(* IEC 61131-3 sources: ST2CPP/examples/projects/syntax_tests, 37 files *)

(* ---- __combined.st ---- *)
(* test_class.st — CLASS 和方法调用测试 *)

CLASS MATH_HELPER
    VAR
        LAST_RESULT : DINT;
        CALL_COUNT  : INT;
    END_VAR

    METHOD ADD : DINT
        VAR_INPUT
            A : DINT;
            B : DINT;
        END_VAR
        LAST_RESULT := A + B;
        CALL_COUNT := CALL_COUNT + 1;
        ADD := LAST_RESULT;
    END_METHOD

    METHOD SUBTRACT : DINT
        VAR_INPUT
            A : DINT;
            B : DINT;
        END_VAR
        LAST_RESULT := A - B;
        CALL_COUNT := CALL_COUNT + 1;
        SUBTRACT := LAST_RESULT;
    END_METHOD

    METHOD GET_COUNT : INT
        GET_COUNT := CALL_COUNT;
    END_METHOD
END_CLASS

PROGRAM TEST_CLASS
    VAR
        Helper      : MATH_HELPER;
        R1          : DINT;
        R2          : DINT;
        Count       : INT;
    END_VAR

    R1 := Helper.ADD(10, 20);
    ASSERT(R1 = 30);

    R2 := Helper.SUBTRACT(50, 15);
    ASSERT(R2 = 35);

    Count := Helper.GET_COUNT();
    ASSERT(Count = 2);

    ASSERT(TRUE);
END_PROGRAM

(* test_class_minimal.st — 最小 CLASS 测试 *)

CLASS BASE_CTRL
    VAR
        BASE_STATE : INT := 0;
    END_VAR

    METHOD GET_VALUE : INT
        GET_VALUE := BASE_STATE;
    END_METHOD
END_CLASS

PROGRAM TEST_MINIMAL
    VAR
        Ctrl : BASE_CTRL;
        R    : INT := 0;
    END_VAR
    R := Ctrl.GET_VALUE();
END_PROGRAM

(* test_class_no_extend.st — CLASS 无继承测试 *)

CLASS MY_CLASS
    VAR
        DATA : INT := 0;
    END_VAR

    METHOD GET_DATA : INT
        GET_DATA := DATA;
    END_METHOD
END_CLASS

PROGRAM TEST_NO_EXTEND
    VAR
        Obj : MY_CLASS;
        R   : INT := 0;
    END_VAR
    R := Obj.GET_DATA();
END_PROGRAM

TYPE MyStruct :
STRUCT
    X : INT;
    Y : INT;
END_STRUCT;
END_TYPE

PROGRAM AT_STRUCT
  VAR_INPUT
    Raw AT %ID0 : MyStruct;
  END_VAR
  VAR_OUTPUT
    Out AT %QD0 : MyStruct;
  END_VAR
  VAR
    LocalX : INT;
  END_VAR
    LocalX := Raw.X;
    Out.Y := Raw.X + 1;
END_PROGRAM

FUNCTION_BLOCK TEST_FB
    VAR_INPUT
        X : INT;
    END_VAR
    VAR_OUTPUT
        Y : INT;
    END_VAR
    VAR
        S : INT := 0;
    END_VAR

    CASE S OF
        0:
            Y := 16#0007;
            IF X > 0 THEN
                S := 1;
            END_IF;
        1:
            Y := 16#000F;
            S := 0;
        ELSE
            Y := 0;
    END_CASE;
END_FUNCTION_BLOCK

PROGRAM IO_TEST
  VAR_INPUT
    BitInput AT %IX1.3 : BOOL;
    ByteInput AT %IB5 : USINT;
    WordInput AT %IW2 : INT;
    DWordInput AT %ID1 : DINT;
  END_VAR
  VAR_OUTPUT
    BitOutput AT %QX0.7 : BOOL;
    ByteOutput AT %QB10 : USINT;
    WordOutput AT %QW3 : INT;
    DWordOutput AT %QD2 : DINT;
  END_VAR
  VAR
    Temp : INT;
    Result : INT;
  END_VAR
    Temp := WordInput + 5;
    IF BitInput THEN
        BitOutput := TRUE;
    ELSE
        BitOutput := FALSE;
    END_IF;
    ByteOutput := ByteInput;
    WordOutput := Temp;
    DWordOutput := DWordInput * 2;
    Result := WordInput * 10;
END_PROGRAM

PROGRAM IO_READBACK
  VAR_INPUT
    Cmd AT %IX0.0 : BOOL;
  END_VAR
  VAR_OUTPUT
    OutVal AT %QW2 : INT;
    OutFlag AT %QX0.1 : BOOL;
  END_VAR
  VAR
    Readback : INT;
    FlagCopy : BOOL;
  END_VAR
    OutVal := 42;
    OutFlag := Cmd;
    Readback := OutVal;
    FlagCopy := OutFlag;
END_PROGRAM

PROGRAM AT_VAR
  VAR
    MyInput AT %IW2 : INT;
    MyOutput AT %QW1 : INT;
    MyFlag AT %QX0.5 : BOOL;
  END_VAR
    MyOutput := MyInput * 2;
    IF MyInput > 100 THEN
        MyFlag := TRUE;
    ELSE
        MyFlag := FALSE;
    END_IF;
END_PROGRAM

(* test_bitwise.st — 测试 Bug 3: AND/OR 对非 BOOL 操作数
 *
 * 问题：VisitAnd_expr 强制要求 BOOL 类型，拒绝 INT 操作数
 * 预期：AND/OR 应支持 ANY_BIT 多态（BYTE/WORD/DWORD/INT 等）
 *       编译器 mapOperator 已将 AND→&, OR→|，只需放宽静态检查
 *)

PROGRAM TEST_BITWISE
    VAR
        A     : INT := 16#FF00;
        B     : INT := 16#0F0F;
        MASK  : INT := 16#00FF;
        AND_R : INT := 0;
        OR_R  : INT := 0;
        XOR_R : INT := 0;
    END_VAR

    AND_R := A AND MASK;
    OR_R  := A OR B;
    XOR_R := A XOR B;

    ASSERT(AND_R = 16#0000);
    ASSERT(OR_R = 16#FF0F);
    ASSERT(XOR_R = 16#F0F0);
END_PROGRAM

FUNCTION_BLOCK MY_FB
    VAR_INPUT X : INT; END_VAR
    VAR_OUTPUT Y : INT; END_VAR
    Y := X + 1;
END_FUNCTION_BLOCK

PROGRAM TEST_FB_ARR
    VAR
        Fbs : ARRAY[0..2] OF MY_FB;
        I : INT;
    END_VAR
    FOR I := 0 TO 2 DO
        Fbs[I](X := I);
    END_FOR;
END_PROGRAM

(* test_fb_output.st — 测试 FB 输出参数 => 在 update 后读回
 *
 * 问题：FB 调用时 => 参数在 update() 后没有从 FB 实例读回
 * 预期：SM(STATUS => MyStatus) 应在 update 后将 FB 的 STATUS 字段读回 MyStatus
 *)

FUNCTION_BLOCK STATE_MACHINE
    VAR_INPUT
        CMD : INT;
    END_VAR
    VAR_OUTPUT
        STATUS : INT;
        DONE   : BOOL;
    END_VAR
    VAR
        MODE : INT := 0;
    END_VAR

    CASE CMD OF
        0:
            MODE := 0;
            STATUS := 0;
            DONE := FALSE;
        1:
            MODE := 1;
            STATUS := 10;
            DONE := TRUE;
        2:
            MODE := 2;
            STATUS := 20;
            DONE := TRUE;
    END_CASE
END_FUNCTION_BLOCK

PROGRAM TEST_FB_OUTPUT
    VAR
        SM       : STATE_MACHINE;
        MyStatus : INT := 0;
        MyDone   : BOOL := FALSE;
    END_VAR

    SM(CMD := 1, STATUS => MyStatus, DONE => MyDone);
    ASSERT(MyStatus = 10);
    ASSERT(MyDone = TRUE);

    SM(CMD := 2, STATUS => MyStatus, DONE => MyDone);
    ASSERT(MyStatus = 20);
    ASSERT(MyDone = TRUE);

    SM(CMD := 0, STATUS => MyStatus, DONE => MyDone);
    ASSERT(MyStatus = 0);
    ASSERT(MyDone = FALSE);
END_PROGRAM

(* test_fc_return.st — 测试 Bug 1: FC 末尾多余 return;
 *
 * 问题：TranslateReturn 对非 void FC 也输出 return; 导致编译报错
 * 预期：非 void FC 应该 return <returnValue>; 而不是 return;
 *)

FUNCTION ADD : DINT
    VAR_INPUT
        A : DINT;
        B : DINT;
    END_VAR
    ADD := A + B;
END_FUNCTION

FUNCTION CLAMP : DINT
    VAR_INPUT
        VAL  : DINT;
        MINV : DINT;
        MAXV : DINT;
    END_VAR
    IF VAL < MINV THEN
        CLAMP := MINV;
    ELSIF VAL > MAXV THEN
        CLAMP := MAXV;
    ELSE
        CLAMP := VAL;
    END_IF
END_FUNCTION

FUNCTION SIMPLE : DINT
    VAR_INPUT
        X : DINT;
    END_VAR
    SIMPLE := X * 2;
    RETURN;
END_FUNCTION

PROGRAM TEST_FC_RETURN
    VAR
        R1 : DINT := 0;
        R2 : DINT := 0;
        R3 : DINT := 0;
    END_VAR
    R1 := ADD(A := 10, B := 20);
    R2 := CLAMP(VAL := -5, MINV := 0, MAXV := 100);
    R3 := SIMPLE(X := 7);

    ASSERT(R1 = 30);
    ASSERT(R2 = 0);
    ASSERT(R3 = 14);
END_PROGRAM

PROGRAM TEST_HEX
    VAR
        X : INT := 0;
        Y : WORD;
    END_VAR
    Y := 16#0007;
    X := 16#FF;
END_PROGRAM

FUNCTION_BLOCK TestFB
    VAR_INPUT LD : BOOL; END_VAR
    VAR_OUTPUT Q : BOOL; END_VAR
END_FUNCTION_BLOCK

PROGRAM main
END_PROGRAM

PROGRAM TEST_ARRAY
    VAR
        JOINT_LIM : ARRAY[0..5, 0..1] OF DINT;
    END_VAR
    JOINT_LIM[0, 0] := -170000;
    JOINT_LIM[0, 1] := 170000;
END_PROGRAM

(* test_not_int.st — AND/OR 位运算测试 *)
(* 注意：当前静态分析器要求 AND/OR 操作数必须为 BOOL *)
(* 此测试验证 BOOL 类型的 AND/OR 生成正确的 & / | *)

PROGRAM TEST_NOT_INT
    VAR
        A       : BOOL;
        B       : BOOL;
        C       : BOOL;
        X       : BOOL := TRUE;
        Y       : BOOL := FALSE;
    END_VAR

    A := TRUE;
    B := FALSE;

    (* AND — 验证生成 & *)
    C := A AND B;
    ASSERT(C = FALSE);

    C := X AND Y;
    ASSERT(C = FALSE);

    C := X AND X;
    ASSERT(C = TRUE);

    (* OR — 验证生成 | *)
    C := A OR B;
    ASSERT(C = TRUE);

    C := Y OR Y;
    ASSERT(C = FALSE);

    C := X OR Y;
    ASSERT(C = TRUE);

    (* NOT — 验证生成 ! *)
    C := NOT X;
    ASSERT(C = FALSE);

    C := NOT Y;
    ASSERT(C = TRUE);

    (* 复合表达式 *)
    C := (X AND Y) OR (X OR Y);
    ASSERT(C = TRUE);

    C := NOT (X AND Y);
    ASSERT(C = TRUE);

    ASSERT(TRUE);
END_PROGRAM

PROGRAM MOTOR_CTRL
  VAR_INPUT
    StartBtn AT %IX0.0 : BOOL;
    StopBtn AT %IX0.1 : BOOL;
    SpeedSensor AT %IW0 : INT;
  END_VAR
  VAR_OUTPUT
    MotorRun AT %QX0.0 : BOOL;
    SpeedOut AT %QW0 : INT;
  END_VAR
  VAR
    TargetSpeed : INT := 1000;
    CurrentSpeed : INT;
    RunLatch : BOOL;
  END_VAR
  VAR RETAIN
    TotalRunTime : DINT;
    ErrorCount : INT;
  END_VAR

  IF StartBtn AND NOT StopBtn THEN
    RunLatch := TRUE;
  END_IF;
  IF StopBtn THEN
    RunLatch := FALSE;
  END_IF;

  MotorRun := RunLatch;

  IF MotorRun THEN
    CurrentSpeed := SpeedSensor;
    SpeedOut := TargetSpeed;
    TotalRunTime := TotalRunTime + 1;
  ELSE
    SpeedOut := 0;
  END_IF;

  IF CurrentSpeed > TargetSpeed * 2 THEN
    ErrorCount := ErrorCount + 1;
  END_IF;
END_PROGRAM

PROGRAM SIMPLE_RETAIN
  VAR
    Counter : INT := 0;
  END_VAR
  VAR RETAIN
    SavedVal : DINT;
  END_VAR

  Counter := Counter + 1;
  SavedVal := SavedVal + Counter;
END_PROGRAM

(* ST2C++ 测试用例 *)

FUNCTION ADD_TEN : INT
    VAR_INPUT
        X : INT;
    END_VAR
    ADD_TEN := X + 10;
END_FUNCTION

PROGRAM P
    VAR
        A : INT := 0;
        B : INT;
    END_VAR

    FOR A := 1 TO 5 BY 1 DO
        B := ADD_TEN(X := A);
    END_FOR
END_PROGRAM

PROGRAM MAIN
  VAR_INPUT
    Start AT %IX0.0 : BOOL;
    Stop AT %IX0.1 : BOOL;
    SpeedRef AT %IW2 : INT;
  END_VAR
  VAR_OUTPUT
    Run AT %QX0.0 : BOOL;
    SpeedOut AT %QW4 : INT;
  END_VAR
  VAR
    Counter : INT;
    Temp AT %IW4 : INT;
    Result AT %QW6 : INT;
  END_VAR
    Counter := Counter + 1;
    IF Start AND NOT Stop THEN
        Run := TRUE;
        SpeedOut := SpeedRef;
    ELSE
        Run := FALSE;
        SpeedOut := 0;
    END_IF;
    Temp := SpeedRef + 10;
    Result := Temp * 2;
END_PROGRAM

(* ---- test_case_hex.st ---- *)
FUNCTION_BLOCK TEST_FB
    VAR_INPUT
        X : INT;
    END_VAR
    VAR_OUTPUT
        Y : INT;
    END_VAR
    VAR
        S : INT := 0;
    END_VAR

    CASE S OF
        0:
            Y := 16#0007;
            IF X > 0 THEN
                S := 1;
            END_IF;
        1:
            Y := 16#000F;
            S := 0;
        ELSE
            Y := 0;
    END_CASE;
END_FUNCTION_BLOCK

(* ---- test_class.st ---- *)
(* test_class.st — CLASS 和方法调用测试 *)

CLASS MATH_HELPER
    VAR
        LAST_RESULT : DINT;
        CALL_COUNT  : INT;
    END_VAR

    METHOD ADD : DINT
        VAR_INPUT
            A : DINT;
            B : DINT;
        END_VAR
        LAST_RESULT := A + B;
        CALL_COUNT := CALL_COUNT + 1;
        ADD := LAST_RESULT;
    END_METHOD

    METHOD SUBTRACT : DINT
        VAR_INPUT
            A : DINT;
            B : DINT;
        END_VAR
        LAST_RESULT := A - B;
        CALL_COUNT := CALL_COUNT + 1;
        SUBTRACT := LAST_RESULT;
    END_METHOD

    METHOD GET_COUNT : INT
        GET_COUNT := CALL_COUNT;
    END_METHOD
END_CLASS

PROGRAM TEST_CLASS
    VAR
        Helper      : MATH_HELPER;
        R1          : DINT;
        R2          : DINT;
        Count       : INT;
    END_VAR

    R1 := Helper.ADD(10, 20);
    ASSERT(R1 = 30);

    R2 := Helper.SUBTRACT(50, 15);
    ASSERT(R2 = 35);

    Count := Helper.GET_COUNT();
    ASSERT(Count = 2);

    ASSERT(TRUE);
END_PROGRAM

(* ---- test_class_minimal.st ---- *)
(* test_class_minimal.st — 最小 CLASS 测试 *)

CLASS BASE_CTRL
    VAR
        BASE_STATE : INT := 0;
    END_VAR

    METHOD GET_VALUE : INT
        GET_VALUE := BASE_STATE;
    END_METHOD
END_CLASS

PROGRAM TEST_MINIMAL
    VAR
        Ctrl : BASE_CTRL;
        R    : INT := 0;
    END_VAR
    R := Ctrl.GET_VALUE();
END_PROGRAM

(* ---- test_class_no_extend.st ---- *)
(* test_class_no_extend.st — CLASS 无继承测试 *)

CLASS MY_CLASS
    VAR
        DATA : INT := 0;
    END_VAR

    METHOD GET_DATA : INT
        GET_DATA := DATA;
    END_METHOD
END_CLASS

PROGRAM TEST_NO_EXTEND
    VAR
        Obj : MY_CLASS;
        R   : INT := 0;
    END_VAR
    R := Obj.GET_DATA();
END_PROGRAM

(* ---- test_class_simple.st ---- *)
(* test_class_simple.st — 简单 CLASS 测试 *)

CLASS MY_CALC
    VAR
        BASE_STATE : INT := 0;
    END_VAR

    METHOD GET_VALUE : INT
        GET_VALUE := INTERNAL;
    END_METHOD
END_CLASS

PROGRAM TEST_SIMPLE
    VAR
        Calc : MY_CALC;
        R    : DINT := 0;
    END_VAR
    R := Calc.GET_VALUE();
END_PROGRAM

(* ---- test_cross_file_type.st ---- *)
(* test_cross_file_type.st — 测试 Bug 2: 跨文件类型解析
 *
 * 问题：多文件编译时 deepFindSymbol 只查 scope chain，不查 PLCTotalSymbolTable
 * 预期：file2.st 能找到 file1.st 中定义的 MY_STRUCT 和 MY_FB
 *)

(* === file1.st 内容 === *)
TYPE
    MY_STRUCT :
    STRUCT
        X : INT;
        Y : DINT;
    END_STRUCT;
END_TYPE

FUNCTION_BLOCK MY_FB
    VAR_INPUT
        CMD : INT;
    END_VAR
    VAR_OUTPUT
        STATE : INT;
    END_VAR
    VAR
        DATA : MY_STRUCT;
    END_VAR

    STATE := CMD;
    DATA.X := CMD;
    DATA.Y := CMD * 10;
END_FUNCTION_BLOCK

(* === file2.st 内容（引用 file1.st 的类型）=== *)
PROGRAM TEST_CROSS_FILE
    VAR
        FB1    : MY_FB;
        RESULT : INT := 0;
        S      : MY_STRUCT;
    END_VAR

    FB1(CMD := 42);
    RESULT := FB1.STATE;
    S.X := 99;

    ASSERT(RESULT = 42);
    ASSERT(S.X = 99);
END_PROGRAM

(* ---- test_fb_array.st ---- *)
FUNCTION_BLOCK MY_FB
    VAR_INPUT X : INT; END_VAR
    VAR_OUTPUT Y : INT; END_VAR
    Y := X + 1;
END_FUNCTION_BLOCK

PROGRAM TEST_FB_ARR
    VAR
        Fbs : ARRAY[0..2] OF MY_FB;
        I : INT;
        R : INT;
    END_VAR
    FOR I := 0 TO 2 DO
        Fbs[I](X := I);
        R := Fbs[I].Y;
    END_FOR;
END_PROGRAM

(* ---- test_fb_array_real.st ---- *)
FUNCTION_BLOCK MY_FB
    VAR_INPUT X : REAL; END_VAR
    VAR_OUTPUT Y : REAL; END_VAR
    Y := X + 1.0;
END_FUNCTION_BLOCK

PROGRAM TEST_FB_ARR
    VAR
        Fbs : ARRAY[0..2] OF MY_FB;
        I : INT;
    END_VAR
    FOR I := 0 TO 2 DO
        Fbs[I](X := 3.14);
    END_FOR;
END_PROGRAM

(* ---- test_fb_array_simple.st ---- *)
FUNCTION_BLOCK MY_FB
    VAR_INPUT X : INT; END_VAR
    VAR_OUTPUT Y : INT; END_VAR
    Y := X + 1;
END_FUNCTION_BLOCK

PROGRAM TEST_FB_ARR
    VAR
        Fbs : ARRAY[0..2] OF MY_FB;
        I : INT;
    END_VAR
    FOR I := 0 TO 2 DO
        Fbs[I](X := I);
    END_FOR;
END_PROGRAM

(* ---- test_fb_init.st ---- *)
TYPE
    JOINT_WAYPOINT :
    STRUCT
        J1      : REAL;
        J2      : REAL;
        SPEED   : REAL;
        DWELL_MS : INT;
    END_STRUCT;
END_TYPE

FUNCTION_BLOCK MY_FB
    VAR_INPUT
        CMD : INT;
    END_VAR
    VAR_OUTPUT
        STATE : INT;
    END_VAR
    VAR
        POS1 : JOINT_WAYPOINT := (J1 := 1.0, J2 := -2.0, SPEED := 10.0, DWELL_MS := 500);
        POS2 : JOINT_WAYPOINT := (J1 := 3.0, J2 := -4.0, SPEED := 20.0, DWELL_MS := 100);
        COUNT : INT := 0;
    END_VAR

    COUNT := COUNT + 1;
END_FUNCTION_BLOCK

PROGRAM TEST_INIT
    VAR
        FB1 : MY_FB;
    END_VAR
END_PROGRAM

(* ---- test_fb_output.st ---- *)
(* test_fb_output.st — 测试 FB 输出参数 => 在 update 后读回
 *
 * 问题：FB 调用时 => 参数在 update() 后没有从 FB 实例读回
 * 预期：SM(STATUS => MyStatus) 应在 update 后将 FB 的 STATUS 字段读回 MyStatus
 *)

FUNCTION_BLOCK STATE_MACHINE
    VAR_INPUT
        CMD : INT;
    END_VAR
    VAR_OUTPUT
        STATUS : INT;
        DONE   : BOOL;
    END_VAR
    VAR
        MODE : INT := 0;
    END_VAR

    CASE CMD OF
        0:
            MODE := 0;
            STATUS := 0;
            DONE := FALSE;
        1:
            MODE := 1;
            STATUS := 10;
            DONE := TRUE;
        2:
            MODE := 2;
            STATUS := 20;
            DONE := TRUE;
    END_CASE
END_FUNCTION_BLOCK

PROGRAM TEST_FB_OUTPUT
    VAR
        SM       : STATE_MACHINE;
        MyStatus : INT := 0;
        MyDone   : BOOL := FALSE;
    END_VAR

    SM(CMD := 1, STATUS => MyStatus, DONE => MyDone);
    ASSERT(MyStatus = 10);
    ASSERT(MyDone = TRUE);

    SM(CMD := 2, STATUS => MyStatus, DONE => MyDone);
    ASSERT(MyStatus = 20);
    ASSERT(MyDone = TRUE);

    SM(CMD := 0, STATUS => MyStatus, DONE => MyDone);
    ASSERT(MyStatus = 0);
    ASSERT(MyDone = FALSE);
END_PROGRAM

(* ---- test_ld.st ---- *)
FUNCTION_BLOCK TestFB
    VAR_INPUT LD : BOOL; END_VAR
    VAR_OUTPUT Q : BOOL; END_VAR
END_FUNCTION_BLOCK

PROGRAM main
END_PROGRAM

(* ---- test_method_output.st ---- *)
(* test_method_output.st — 测试 Bug 5: CLASS 方法输出参数 =>
 *
 * 问题：调用端把 => 参数原样 dump 成无效 C++（STATE_OUT => myVar）
 * 预期：=> 参数应翻译为 C++ 引用传递，调用后写回变量
 * 注意：INTERNAL 是保留字，不能用作变量名
 *)

CLASS MY_CALC
    VAR
        ACCUM : DINT := 0;
    END_VAR

    METHOD ADD_AND_REPORT : DINT
        VAR_INPUT
            VALUE : DINT;
        END_VAR
        VAR_OUTPUT
            REPORT : DINT;
        END_VAR
        ACCUM := ACCUM + VALUE;
        REPORT := ACCUM;
        ADD_AND_REPORT := ACCUM;
    END_METHOD
END_CLASS

PROGRAM TEST_METHOD_OUTPUT
    VAR
        Calc     : MY_CALC;
        MyReport : DINT := 0;
        Result   : DINT := 0;
    END_VAR

    Result := Calc.ADD_AND_REPORT(VALUE := 10, REPORT => MyReport);
    ASSERT(Result = 10);
    ASSERT(MyReport = 10);

    Result := Calc.ADD_AND_REPORT(VALUE := 20, REPORT => MyReport);
    ASSERT(Result = 30);
    ASSERT(MyReport = 30);
END_PROGRAM

(* ---- test_super.st ---- *)
(* test_super.st — SUPER:: 调用测试 *)

CLASS BASE_CALC
    VAR
        BASE_VALUE : DINT;
    END_VAR

    METHOD INIT_BASE
        VAR_INPUT
            VAL : DINT;
        END_VAR
        BASE_VALUE := VAL;
    END_METHOD

    METHOD GET_VALUE : DINT
        GET_VALUE := BASE_VALUE;
    END_METHOD
END_CLASS

CLASS EXTEND_CALC EXTENDS BASE_CALC
    VAR
        EXT_VALUE : DINT;
    END_VAR

    METHOD INIT_EXT
        VAR_INPUT
            BASE_VAL : DINT;
            EXT_VAL  : DINT;
        END_VAR
        SUPER.INIT_BASE();
        EXT_VALUE := EXT_VAL;
    END_METHOD

    METHOD GET_TOTAL : DINT
        GET_TOTAL := SUPER.GET_VALUE() + EXT_VALUE;
    END_METHOD
END_CLASS

PROGRAM TEST_SUPER
    VAR
        Calc    : EXTEND_CALC;
        R1      : DINT;
    END_VAR

    Calc.INIT_EXT();
    R1 := Calc.GET_TOTAL();
    ASSERT(TRUE);
END_PROGRAM

(* ---- test_super_call.st ---- *)
(* test_super_call.st — 测试 Bug 4: SUPER:: 调用
 *
 * 问题：SUPER.MethodName() 只输出注释，不生成实际父类调用
 * 预期：SUPER. 应翻译为 ParentClass::MethodName(this, ...) 的 C++ 调用
 * 注意：ST 标准语法是 SUPER.method() 而非 SUPER::method()
 *)

CLASS BASE_CTRL
    VAR
        BASE_STATE : INT := 0;
    END_VAR

    METHOD INIT_BASE : INT
        BASE_STATE := 1;
        INIT_BASE := BASE_STATE;
    END_METHOD
END_CLASS

CLASS CHILD_CTRL EXTENDS BASE_CTRL
    VAR
        CHILD_DATA : INT := 0;
    END_VAR

    METHOD INIT_CHILD : INT
        SUPER.INIT_BASE();
        CHILD_DATA := 42;
        INIT_CHILD := CHILD_DATA;
    END_METHOD
END_CLASS

PROGRAM TEST_SUPER
    VAR
        Child : CHILD_CTRL;
        R     : INT := 0;
    END_VAR

    R := Child.INIT_CHILD();
    ASSERT(R = 42);
END_PROGRAM

(* ---- test_to.st ---- *)
FUNCTION_BLOCK TestFB
    VAR_INPUT TO : BOOL; END_VAR
    VAR_OUTPUT Q : BOOL; END_VAR
END_FUNCTION_BLOCK

PROGRAM main
END_PROGRAM

(* ---- test_tricky.st ---- *)
(*
 * test_tricky.st — 刁钻综合测试
 *
 * 覆盖:
 *   1. ENUM + CASE 分支 (语法: TYPE NAME : (VAL1, VAL2); END_TYPE)
 *   2. 嵌套 FOR + 结构体数组
 *   3. WHILE/REPEAT 循环
 *   4. 多返回路径函数
 *   5. 函数调用函数
 *   6. 混合类型运算 (INT/DINT/REAL)
 *   7. 复杂布尔表达式 (AND/OR/NOT)
 *   8. STRING 拼接 (PRINT)
 *)

TYPE
    DIRECTION : (NORTH, EAST, SOUTH, WEST);
END_TYPE

TYPE
    MATRIX_ROW :
    STRUCT
        VALUES : ARRAY[0..3] OF INT;
        TAG    : INT;
    END_STRUCT;
END_TYPE

FUNCTION DOUBLE_IT : DINT
    VAR_INPUT
        X : INT;
    END_VAR
    DOUBLE_IT := X * 2;
END_FUNCTION

FUNCTION CLAMP : DINT
    VAR_INPUT
        VAL  : DINT;
        MINV : DINT;
        MAXV : DINT;
    END_VAR
    IF VAL < MINV THEN
        CLAMP := MINV;
    ELSIF VAL > MAXV THEN
        CLAMP := MAXV;
    ELSE
        CLAMP := VAL;
    END_IF
END_FUNCTION

FUNCTION WRAP_ANGLE : INT
    VAR_INPUT
        ANGLE : INT;
    END_VAR
    WHILE ANGLE < 0 DO
        ANGLE := ANGLE + 360;
    END_WHILE
    WHILE ANGLE >= 360 DO
        ANGLE := ANGLE - 360;
    END_WHILE
    WRAP_ANGLE := ANGLE;
END_FUNCTION

FUNCTION AVERAGE : REAL
    VAR_INPUT
        A : REAL;
        B : REAL;
    END_VAR
    AVERAGE := (A + B) / 2.0;
END_FUNCTION

FUNCTION_BLOCK STATE_MACHINE
    VAR_INPUT
        CMD      : INT;
        POSITION : DINT;
    END_VAR
    VAR_OUTPUT
        DIR      : DIRECTION;
        SPEED    : INT;
        FAULT    : BOOL;
    END_VAR
    VAR
        MODE     : INT := 0;
        ACCUM    : DINT := 0;
        RUNNING  : BOOL := FALSE;
        RETRY    : INT := 0;
    END_VAR

    FAULT := FALSE;
    RUNNING := TRUE;

    CASE CMD OF
        0:
            MODE := 0;
            ACCUM := 0;
            SPEED := 0;
            DIR := DIRECTION#NORTH;
            RUNNING := FALSE;
        1:
            MODE := 10;
            ACCUM := 0;
            DIR := DIRECTION#EAST;
        2:
            MODE := 20;
            ACCUM := 0;
            DIR := DIRECTION#WEST;
        3:
            MODE := 30;
            DIR := DIRECTION#SOUTH;
        10:
            MODE := 0;
            FAULT := TRUE;
        ELSE
            MODE := 99;
            FAULT := TRUE;
    END_CASE

    IF RUNNING THEN
        CASE MODE OF
            10:
                ACCUM := ACCUM + POSITION;
                IF ACCUM >= 1000 THEN
                    MODE := 11;
                END_IF
            20:
                ACCUM := ACCUM - POSITION;
                IF ACCUM <= -1000 THEN
                    MODE := 21;
                END_IF
            30:
                SPEED := 0;
                RETRY := RETRY + 1;
                IF RETRY >= 3 THEN
                    MODE := 31;
                END_IF
            11, 21, 31:
                SPEED := 0;
                RUNNING := FALSE;
        END_CASE
    END_IF
END_FUNCTION_BLOCK

PROGRAM TRICKY_MAIN
    VAR
        MATRIX    : ARRAY[0..2] OF MATRIX_ROW;
        I         : INT := 0;
        J         : INT := 0;
        TOTAL     : DINT := 0;
        COUNT     : DINT := 0;
        VAL       : INT := -450;
        WRAPPED   : INT := 0;
        AVG       : REAL := 0.0;
        CLAMPED   : DINT := 0;
        CLAMPED2  : DINT := 0;
        SM        : STATE_MACHINE;
        PHASE     : INT := 0;
        FLAG      : BOOL := FALSE;
        RESULT_ARR : ARRAY[0..5] OF DINT;
        K         : INT := 0;
        ARR_VAL   : DINT := 0;
    END_VAR

    PRINT("=== TRICKY TEST START ===");

    (* 1. 嵌套 FOR + STRUCT 数组赋值 *)
    FOR I := 0 TO 2 BY 1 DO
        MATRIX[I].TAG := I * 100;
        FOR J := 0 TO 3 BY 1 DO
            MATRIX[I].VALUES[J] := (I * 10) + J;
            TOTAL := TOTAL + MATRIX[I].VALUES[J];
        END_FOR
    END_FOR

    PRINT("TOTAL = " + TOTAL);

    (* 2. WHILE 取模 (角度归约) *)
    WRAPPED := WRAP_ANGLE(ANGLE := VAL);
    PRINT("WRAPPED = " + WRAPPED);

    (* 3. 函数调用函数 (浮点) *)
    AVG := AVERAGE(A := 10.5, B := 20.5);
    PRINT("AVG = " + AVG);

    (* 4. 多返回路径 (CLAMP) *)
    CLAMPED := CLAMP(VAL := -100, MINV := 0, MAXV := 50);
    PRINT("CLAMPED = " + CLAMPED);
    CLAMPED2 := CLAMP(VAL := 999, MINV := 0, MAXV := 100);
    PRINT("CLAMPED2 = " + CLAMPED2);

    (* 5. ENUM + CASE 状态机 *)
    PHASE := 1;
    SM(CMD := PHASE, POSITION := 500);
    PHASE := 2;
    SM(CMD := PHASE, POSITION := 1200);
    PHASE := 3;
    SM(CMD := PHASE, POSITION := -800);

    (* 6. REPEAT 循环 *)
    K := 0;
    REPEAT
        RESULT_ARR[K] := DOUBLE_IT(X := K * 10);
        K := K + 1;
    UNTIL K >= 6
    END_REPEAT

    ARR_VAL := 42;
    PRINT("RESULT_ARR[3] = " + ARR_VAL);

    (* 7. 复杂布尔表达式 *)
    FLAG := (I >= 2) AND (TOTAL > 0) OR (WRAPPED <> 270);
    IF FLAG AND NOT (CLAMPED < 0) THEN
        PRINT("FLAG IS TRUE");
    END_IF

    (* 8. WHILE 模拟 BREAK *)
    COUNT := 0;
    WHILE COUNT < 10 DO
        COUNT := COUNT + 1;
        IF COUNT = 5 THEN
            COUNT := 10;
        END_IF
    END_WHILE
    PRINT("COUNT = " + COUNT);

    (* 9. ASSERT 综合验证 *)
    ASSERT(TOTAL = 66);
    ASSERT(WRAPPED = 270);
    ASSERT(CLAMPED = 50);
    ASSERT(AVG > 15.0);
    ASSERT(MATRIX[0].TAG = 0);
    ASSERT(MATRIX[2].VALUES[3] = 23);
    ASSERT(K >= 6);
    ASSERT(NOT FLAG);

    PRINT("=== TRICKY TEST PASS ===");
END_PROGRAM

(* ---- test_tricky_mini.st ---- *)
TYPE
    DIRECTION : (NORTH, EAST, SOUTH, WEST);
END_TYPE

FUNCTION_BLOCK MINI
    VAR_OUTPUT
        DIR : INT;
    END_VAR
    VAR
        STP : INT := 0;
    END_VAR
    DIR := 42;
END_FUNCTION_BLOCK

PROGRAM MAIN
    VAR
        M : MINI;
    END_VAR
    M();
END_PROGRAM

(* ---- demo_at.st ---- *)
PROGRAM DEMO
  VAR_INPUT
    Start AT %IX0.0 : BOOL;
    Stop AT %IX0.1 : BOOL;
    SpeedRef AT %IW2 : INT;
  END_VAR
  VAR_OUTPUT
    Run AT %QX0.0 : BOOL;
    SpeedOut AT %QW4 : INT;
  END_VAR
  VAR
    Counter : INT;
    Temp AT %IW6 : INT;
  END_VAR
    Counter := Counter + 1;
    IF Start AND NOT Stop THEN
        Run := TRUE;
        SpeedOut := SpeedRef;
    ELSE
        Run := FALSE;
        SpeedOut := 0;
    END_IF;
    SpeedOut := SpeedRef + Temp;
END_PROGRAM

(* ---- test.st ---- *)
(* ST2C++ 测试用例 *)

FUNCTION ADD_TEN : INT
    VAR_INPUT
        X : INT;
    END_VAR
    ADD_TEN := X + 10;
END_FUNCTION

PROGRAM P
    VAR
        A : INT := 0;
        B : INT;
    END_VAR

    FOR A := 1 TO 5 BY 1 DO
        B := ADD_TEN(X := A);
    END_FOR
END_PROGRAM

(* ---- test_arr_struct.st ---- *)
TYPE
    MY_POINT :
    STRUCT
        X : INT;
        Y : INT;
    END_STRUCT;
END_TYPE

PROGRAM MAIN
    VAR
        P_ARR : ARRAY[0..4] OF MY_POINT;
        I : INT := 0;
        SUM_X : INT := 0;
    END_VAR

    FOR I := 0 TO 4 BY 1 DO
        P_ARR[I].X := I * 10;
        P_ARR[I].Y := I * 20;
    END_FOR

    SUM_X := P_ARR[0].X + P_ARR[1].X;
END_PROGRAM

(* ---- test_at.st ---- *)
PROGRAM MAIN
  VAR_INPUT
    Start AT %IX0.0 : BOOL;
    Stop AT %IX0.1 : BOOL;
    SpeedRef AT %IW2 : INT;
  END_VAR
  VAR_OUTPUT
    Run AT %QX0.0 : BOOL;
    SpeedOut AT %QW4 : INT;
  END_VAR
  VAR
    Counter : INT;
    Temp AT %IW4 : INT;
    Result AT %QW6 : INT;
  END_VAR
    Counter := Counter + 1;
    IF Start AND NOT Stop THEN
        Run := TRUE;
        SpeedOut := SpeedRef;
    ELSE
        Run := FALSE;
        SpeedOut := 0;
    END_IF;
    Temp := SpeedRef + 10;
    Result := Temp * 2;
END_PROGRAM

(* ---- test_at_full.st ---- *)
PROGRAM IO_TEST
  VAR_INPUT
    BitInput AT %IX1.3 : BOOL;
    ByteInput AT %IB5 : USINT;
    WordInput AT %IW2 : INT;
    DWordInput AT %ID1 : DINT;
  END_VAR
  VAR_OUTPUT
    BitOutput AT %QX0.7 : BOOL;
    ByteOutput AT %QB10 : USINT;
    WordOutput AT %QW3 : INT;
    DWordOutput AT %QD2 : DINT;
  END_VAR
  VAR
    Temp : INT;
    Result : INT;
  END_VAR
    Temp := WordInput + 5;
    IF BitInput THEN
        BitOutput := TRUE;
    ELSE
        BitOutput := FALSE;
    END_IF;
    ByteOutput := ByteInput;
    WordOutput := Temp;
    DWordOutput := DWordInput * 2;
    Result := WordInput * 10;
END_PROGRAM

(* ---- test_at_output_read.st ---- *)
PROGRAM IO_READBACK
  VAR_INPUT
    Cmd AT %IX0.0 : BOOL;
  END_VAR
  VAR_OUTPUT
    OutVal AT %QW2 : INT;
    OutFlag AT %QX0.1 : BOOL;
  END_VAR
  VAR
    Readback : INT;
    FlagCopy : BOOL;
  END_VAR
    OutVal := 42;
    OutFlag := Cmd;
    Readback := OutVal;
    FlagCopy := OutFlag;
END_PROGRAM

(* ---- test_at_struct.st ---- *)
TYPE MyStruct :
STRUCT
    X : INT;
    Y : INT;
END_STRUCT;
END_TYPE

PROGRAM AT_STRUCT
  VAR_INPUT
    Raw AT %ID0 : MyStruct;
  END_VAR
  VAR_OUTPUT
    Out AT %QD0 : MyStruct;
  END_VAR
  VAR
    LocalX : INT;
  END_VAR
    LocalX := Raw.X;
    Out.Y := Raw.X + 1;
END_PROGRAM

(* ---- test_at_var.st ---- *)
PROGRAM AT_VAR
  VAR
    MyInput AT %IW2 : INT;
    MyOutput AT %QW1 : INT;
    MyFlag AT %QX0.5 : BOOL;
  END_VAR
    MyOutput := MyInput * 2;
    IF MyInput > 100 THEN
        MyFlag := TRUE;
    ELSE
        MyFlag := FALSE;
    END_IF;
END_PROGRAM

(* ---- test_bitwise.st ---- *)
(* test_bitwise.st — 测试 Bug 3: AND/OR 对非 BOOL 操作数
 *
 * 问题：VisitAnd_expr 强制要求 BOOL 类型，拒绝 INT 操作数
 * 预期：AND/OR 应支持 ANY_BIT 多态（BYTE/WORD/DWORD/INT 等）
 *       编译器 mapOperator 已将 AND→&, OR→|，只需放宽静态检查
 *)

PROGRAM TEST_BITWISE
    VAR
        A     : INT := 16#FF00;
        B     : INT := 16#0F0F;
        MASK  : INT := 16#00FF;
        AND_R : INT := 0;
        OR_R  : INT := 0;
        XOR_R : INT := 0;
    END_VAR

    AND_R := A AND MASK;
    OR_R  := A OR B;
    XOR_R := A XOR B;

    ASSERT(AND_R = 16#0000);
    ASSERT(OR_R = 16#FF0F);
    ASSERT(XOR_R = 16#F0F0);
END_PROGRAM

(* ---- test_fc_return.st ---- *)
(* test_fc_return.st — 测试 Bug 1: FC 末尾多余 return;
 *
 * 问题：TranslateReturn 对非 void FC 也输出 return; 导致编译报错
 * 预期：非 void FC 应该 return <returnValue>; 而不是 return;
 *)

FUNCTION ADD : DINT
    VAR_INPUT
        A : DINT;
        B : DINT;
    END_VAR
    ADD := A + B;
END_FUNCTION

FUNCTION CLAMP : DINT
    VAR_INPUT
        VAL  : DINT;
        MINV : DINT;
        MAXV : DINT;
    END_VAR
    IF VAL < MINV THEN
        CLAMP := MINV;
    ELSIF VAL > MAXV THEN
        CLAMP := MAXV;
    ELSE
        CLAMP := VAL;
    END_IF
END_FUNCTION

FUNCTION SIMPLE : DINT
    VAR_INPUT
        X : DINT;
    END_VAR
    SIMPLE := X * 2;
    RETURN;
END_FUNCTION

PROGRAM TEST_FC_RETURN
    VAR
        R1 : DINT := 0;
        R2 : DINT := 0;
        R3 : DINT := 0;
    END_VAR
    R1 := ADD(A := 10, B := 20);
    R2 := CLAMP(VAL := -5, MINV := 0, MAXV := 100);
    R3 := SIMPLE(X := 7);

    ASSERT(R1 = 30);
    ASSERT(R2 = 0);
    ASSERT(R3 = 14);
END_PROGRAM

(* ---- test_hex.st ---- *)
PROGRAM TEST_HEX
    VAR
        X : INT := 0;
        Y : WORD;
    END_VAR
    Y := 16#0007;
    X := 16#FF;
END_PROGRAM

(* ---- test_multidim.st ---- *)
PROGRAM TEST_ARRAY
    VAR
        JOINT_LIM : ARRAY[0..5, 0..1] OF DINT;
    END_VAR
    JOINT_LIM[0, 0] := -170000;
    JOINT_LIM[0, 1] := 170000;
END_PROGRAM

(* ---- test_not_int.st ---- *)
(* test_not_int.st — AND/OR 位运算测试 *)
(* 注意：当前静态分析器要求 AND/OR 操作数必须为 BOOL *)
(* 此测试验证 BOOL 类型的 AND/OR 生成正确的 & / | *)

PROGRAM TEST_NOT_INT
    VAR
        A       : BOOL;
        B       : BOOL;
        C       : BOOL;
        X       : BOOL := TRUE;
        Y       : BOOL := FALSE;
    END_VAR

    A := TRUE;
    B := FALSE;

    (* AND — 验证生成 & *)
    C := A AND B;
    ASSERT(C = FALSE);

    C := X AND Y;
    ASSERT(C = FALSE);

    C := X AND X;
    ASSERT(C = TRUE);

    (* OR — 验证生成 | *)
    C := A OR B;
    ASSERT(C = TRUE);

    C := Y OR Y;
    ASSERT(C = FALSE);

    C := X OR Y;
    ASSERT(C = TRUE);

    (* NOT — 验证生成 ! *)
    C := NOT X;
    ASSERT(C = FALSE);

    C := NOT Y;
    ASSERT(C = TRUE);

    (* 复合表达式 *)
    C := (X AND Y) OR (X OR Y);
    ASSERT(C = TRUE);

    C := NOT (X AND Y);
    ASSERT(C = TRUE);

    ASSERT(TRUE);
END_PROGRAM

(* ---- test_pre_post.st ---- *)
PROGRAM MOTOR_CTRL
  VAR_INPUT
    StartBtn AT %IX0.0 : BOOL;
    StopBtn AT %IX0.1 : BOOL;
    SpeedSensor AT %IW0 : INT;
  END_VAR
  VAR_OUTPUT
    MotorRun AT %QX0.0 : BOOL;
    SpeedOut AT %QW0 : INT;
  END_VAR
  VAR
    TargetSpeed : INT := 1000;
    CurrentSpeed : INT;
    RunLatch : BOOL;
  END_VAR
  VAR RETAIN
    TotalRunTime : DINT;
    ErrorCount : INT;
  END_VAR

  IF StartBtn AND NOT StopBtn THEN
    RunLatch := TRUE;
  END_IF;
  IF StopBtn THEN
    RunLatch := FALSE;
  END_IF;

  MotorRun := RunLatch;

  IF MotorRun THEN
    CurrentSpeed := SpeedSensor;
    SpeedOut := TargetSpeed;
    TotalRunTime := TotalRunTime + 1;
  ELSE
    SpeedOut := 0;
  END_IF;

  IF CurrentSpeed > TargetSpeed * 2 THEN
    ErrorCount := ErrorCount + 1;
  END_IF;
END_PROGRAM

(* ---- test_retain_simple.st ---- *)
PROGRAM SIMPLE_RETAIN
  VAR
    Counter : INT := 0;
  END_VAR
  VAR RETAIN
    SavedVal : DINT;
  END_VAR

  Counter := Counter + 1;
  SavedVal := SavedVal + Counter;
END_PROGRAM

(* ---- test_std_fb.st ---- *)
PROGRAM main
  VAR myTimer : TON; END_VAR
  myTimer(IN:=TRUE, PT:=T#500ms);
END_PROGRAM

(* ---- test_struct.st ---- *)
TYPE
    MY_POINT :
    STRUCT
        X : INT;
        Y : INT;
    END_STRUCT;
END_TYPE

PROGRAM MAIN
    VAR
        P : MY_POINT;
        SUM : INT := 0;
    END_VAR

    P.X := 10;
    P.Y := 20;
    SUM := P.X + P.Y;
END_PROGRAM

(* ---- traffic_light.st ---- *)
(* traffic_light.st — 十字路口交通灯控制 *)

PROGRAM TRAFFIC_LIGHT
    VAR
        phase       : INT := 1;
        tick_count  : DINT := 0;
        green_ticks : DINT := 3000;
        yellow_ticks: DINT := 500;
        clear_ticks : DINT := 200;
        ns_r        : BOOL := TRUE;
        ns_y        : BOOL := FALSE;
        ns_g        : BOOL := FALSE;
        ew_r        : BOOL := TRUE;
        ew_y        : BOOL := FALSE;
        ew_g        : BOOL := FALSE;
    END_VAR

    tick_count := tick_count + 1;

    IF phase = 1 AND tick_count >= green_ticks THEN
        tick_count := 0;
        phase := 2;
    ELSIF phase = 2 AND tick_count >= yellow_ticks THEN
        tick_count := 0;
        phase := 3;
    ELSIF phase = 3 AND tick_count >= clear_ticks THEN
        tick_count := 0;
        phase := 4;
    ELSIF phase = 4 AND tick_count >= green_ticks THEN
        tick_count := 0;
        phase := 5;
    ELSIF phase = 5 AND tick_count >= yellow_ticks THEN
        tick_count := 0;
        phase := 6;
    ELSIF phase = 6 AND tick_count >= clear_ticks THEN
        tick_count := 0;
        phase := 1;
    END_IF;

    ns_r := FALSE;
    ns_y := FALSE;
    ns_g := FALSE;
    ew_r := FALSE;
    ew_y := FALSE;
    ew_g := FALSE;

    IF phase = 1 THEN
        ns_g := TRUE;
        ew_r := TRUE;
    ELSIF phase = 2 THEN
        ns_y := TRUE;
        ew_r := TRUE;
    ELSIF phase = 3 THEN
        ns_r := TRUE;
        ew_r := TRUE;
    ELSIF phase = 4 THEN
        ns_r := TRUE;
        ew_g := TRUE;
    ELSIF phase = 5 THEN
        ns_r := TRUE;
        ew_y := TRUE;
    ELSE
        ns_r := TRUE;
        ew_r := TRUE;
    END_IF;

END_PROGRAM
